Fanuc KAREL source: kx00006.KL

-- PROVISIONAL review KL for V1013-1; original PC SHA256 92144a005acca1b5e47958b75c95c13f03cd0b1f90a1ea8597343a755733e651
-- Incomplete behavior may be omitted. Consult companion uncertainty JSON. Do not deploy.
PROGRAM KX00006
%NOLOCKGROUP
VAR
  I : INTEGER
  J : INTEGER
  B : BOOLEAN
  F : FILE
  S : STRING[80]
-- UNRESOLVED_DECL P type=000102
BEGIN
  -- UNRESOLVED_PC offsets 5-13; opcodes 9D,2E,0F
  -- UNRESOLVED_PC offsets 18-22; opcodes 7F
END KX00006
